(* IEC 61131-3 sources: cds-text-sync/products/codesys-agent/tests/Cts.Agent.Core.Tests/Golden/ExportFixture/folder-case, 1 file *)

(* ---- I_LiveTmp.st ---- *)
INTERFACE I_LiveTmp
END_INTERFACE

METHOD M_LiveTmp : BOOL
VAR_INPUT
	x : BOOL;
END_VAR
END_METHOD
